(* IEC 61131-3 sources: volt/packages/volt-lsp-iec/test-corpus/bakon-nano/Device/Plc Logic/Application/Library Manager/CmpSchedule, 15 files *)

(* ---- SCHEDGETCURRENTTASK.pou ---- *)
FUNCTION SCHEDGETCURRENTTASK : RTS_IEC_HANDLE
VAR_INPUT
	PRESULT : POINTER TO RTS_IEC_RESULT;
END_VAR
END_FUNCTION

(* ---- SCHEDGETNUMOFTASKS.pou ---- *)
FUNCTION SCHEDGETNUMOFTASKS : DINT
VAR_INPUT
	PAPP : POINTER TO APPLICATION;
	PRESULT : POINTER TO RTS_IEC_RESULT;
END_VAR
END_FUNCTION

(* ---- SCHEDGETPROCESSORLOAD.pou ---- *)
FUNCTION SCHEDGETPROCESSORLOAD : UDINT
VAR_INPUT
	PRESULT : POINTER TO RTS_IEC_RESULT;
END_VAR
END_FUNCTION

(* ---- SCHEDGETTASKEVENTBYHANDLE.pou ---- *)
FUNCTION SCHEDGETTASKEVENTBYHANDLE : RTS_IEC_HANDLE
VAR_INPUT
	HSCHEDTASK : RTS_IEC_HANDLE;
	PRESULT : POINTER TO RTS_IEC_RESULT;
END_VAR
END_FUNCTION

(* ---- SCHEDGETTASKHANDLEBYINDEX.pou ---- *)
FUNCTION SCHEDGETTASKHANDLEBYINDEX : RTS_IEC_HANDLE
VAR_INPUT
	PAPP : POINTER TO APPLICATION;
	NINDEX : DINT;
	PRESULT : POINTER TO RTS_IEC_RESULT;
END_VAR
END_FUNCTION

(* ---- SCHEDGETTASKHANDLEBYNAME.pou ---- *)
FUNCTION SCHEDGETTASKHANDLEBYNAME : RTS_IEC_HANDLE
VAR_INPUT
	PRESULT : POINTER TO RTS_IEC_RESULT;
END_VAR
VAR_IN_OUT
	PSZTASKNAME : STRING;
END_VAR
END_FUNCTION

(* ---- SCHEDGETTASKINTERVAL.pou ---- *)
FUNCTION SCHEDGETTASKINTERVAL : RTS_IEC_RESULT
VAR_INPUT
	HSCHEDTASK : RTS_IEC_HANDLE;
END_VAR
VAR_IN_OUT
	PULINTERVAL : UDINT;
END_VAR
END_FUNCTION

(* ---- SCHEDPOSTEXTERNALEVENT.pou ---- *)
FUNCTION SCHEDPOSTEXTERNALEVENT : RTS_IEC_RESULT
VAR_INPUT
	HEXTEVENT : RTS_IEC_HANDLE;
END_VAR
END_FUNCTION

(* ---- SCHEDREGISTEREXTERNALEVENT.pou ---- *)
FUNCTION SCHEDREGISTEREXTERNALEVENT : RTS_IEC_HANDLE
VAR_INPUT
	PSZEXTEVENTNAME : REFERENCE TO STRING;
	PRESULT : POINTER TO RTS_IEC_RESULT;
END_VAR
END_FUNCTION

(* ---- SCHEDSETTASKINTERVAL.pou ---- *)
FUNCTION SCHEDSETTASKINTERVAL : RTS_IEC_RESULT
VAR_INPUT
	HSCHEDTASK : RTS_IEC_HANDLE;
	ULINTERVAL : UDINT;
END_VAR
END_FUNCTION

(* ---- SCHEDTASKRESUME.pou ---- *)
FUNCTION SCHEDTASKRESUME : SysTypes.RTS_IEC_RESULT
VAR_INPUT
	HSCHEDTASK : SysTypes.RTS_IEC_HANDLE;
END_VAR
END_FUNCTION

(* ---- SCHEDTASKSUSPEND.pou ---- *)
FUNCTION SCHEDTASKSUSPEND : SysTypes.RTS_IEC_RESULT
VAR_INPUT
	HSCHEDTASK : SysTypes.RTS_IEC_HANDLE;
END_VAR
END_FUNCTION

(* ---- SCHEDUNREGISTEREXTERNALEVENT.pou ---- *)
FUNCTION SCHEDUNREGISTEREXTERNALEVENT : RTS_IEC_RESULT
VAR_INPUT
	HEXTEVENT : RTS_IEC_HANDLE;
END_VAR
END_FUNCTION

(* ---- SCHEDWAITBUSY.pou ---- *)
FUNCTION SCHEDWAITBUSY : RTS_IEC_RESULT
VAR_IN_OUT
	PTSLEEPUS : SYSTIME;
END_VAR
END_FUNCTION

(* ---- SCHEDWAITSLEEP.pou ---- *)
FUNCTION SCHEDWAITSLEEP : RTS_IEC_RESULT
VAR_IN_OUT
	PTSLEEPUS : SYSTIME;
END_VAR
END_FUNCTION
